TYPE "FRK_Document_D011"
VERSION : 0.1
   STRUCT
      SchemaVersion { ExternalAccessible := 'False'; ExternalVisible := 'False'; ExternalWritable := 'False'} : UInt;
      Scope { ExternalAccessible := 'False'; ExternalVisible := 'False'; ExternalWritable := 'False'} : String[80];
      Image { ExternalAccessible := 'False'; ExternalVisible := 'False'; ExternalWritable := 'False'} : "ST_LineImage";
   END_STRUCT;

END_TYPE

